FUNCTION_BLOCK IO_RouteDI (* Picks the way an IO block reaches its signal from the Address (a Pi line, a local IO handle, Modbus or simulated) and passes values through that way only. Technical: Backend router for IO_DI; Address: 'gpio[chip:line(:pull_up|:pull_down)(:active_low)]' or 'pwm[chip:channel:period_ns]' a Raspberry Pi's line, set up here; 'modbus[...]' a Modbus CLIENT ID; 'sim' simulated; another name a local IO handle set up elsewhere (IX/QX PARAMS); empty: not connected (QO = FALSE) *)
  (* Standard: 61499-2 *)
  (* Version 0.1, 2026-09-28, Project contributors, AAU Smart Production Lab *)
  PACKAGE modlib;
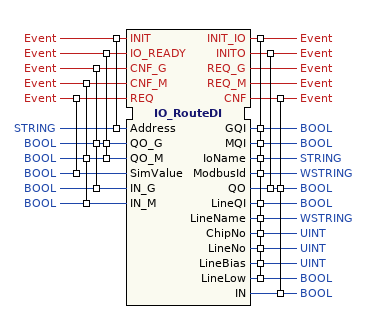
  EVENT_INPUT
    INIT WITH Address; (* Work out from Address how the point is reached *)
    IO_READY WITH QO_G, QO_M; (* The line, the local IO block and the Modbus client are initialised *)
    CNF_G WITH QO_G, IN_G; (* The local IO block answered *)
    CNF_M WITH QO_M, IN_M; (* The Modbus client answered *)
    REQ WITH SimValue; (* Access the point *)
  END_EVENT
  EVENT_OUTPUT
    INIT_IO WITH GQI, MQI, IoName, ModbusId, LineQI, LineName, ChipNo, LineNo, LineBias, LineLow; (* Set up the line, the local IO block and the Modbus client (each only if it is the way) *)
    INITO WITH QO; (* Initialised: QO says whether the point is reachable *)
    REQ_G; (* Access the point through the local IO block (IX/QX/IW/QW) *)
    REQ_M; (* Access the point through the Modbus client *)
    CNF WITH QO, IN; (* Done: QO says whether it worked *)
  END_EVENT
  VAR_INPUT
    Address : STRING; (* Where the point is: 'gpio[chip:line(:pull_up|:pull_down)(:active_low)]', 'pwm[chip:channel:period_ns]', 'modbus[...]', 'sim', or an IO handle's name; empty: not connected *)
    QO_G : BOOL; (* The local IO block works *)
    QO_M : BOOL; (* The Modbus client works *)
    SimValue : BOOL; (* The value read when the address is 'sim' *)
    IN_G : BOOL; (* The raw value read through the local IO block *)
    IN_M : BOOL; (* The raw value read through Modbus *)
  END_VAR
  VAR_OUTPUT
    GQI : BOOL; (* Use the local IO block *)
    MQI : BOOL; (* Use the Modbus client *)
    IoName : STRING; (* The local IO handle's name (PARAMS of IX/QX/IW/QW) *)
    ModbusId : WSTRING; (* The Modbus CLIENT's ID *)
    QO : BOOL; (* The point is reachable, the last access worked *)
    LineQI : BOOL; (* Set up a Raspberry Pi line here (a gpio[...] or pwm[...] address) *)
    LineName : WSTRING; (* The name the line is registered under (the address) *)
    ChipNo : UINT; (* The GPIO or PWM chip's number *)
    LineNo : UINT; (* The GPIO line's or PWM channel's number *)
    LineBias : UINT; (* GPIO bias: 0 none, 2 pull-up, 3 pull-down (FORTE 3.3.0's numbering) *)
    LineLow : BOOL; (* The line is active low *)
    IN : BOOL; (* The value read (an analog one scaled) *)
  END_VAR
  VAR
    Backend : USINT;
  END_VAR
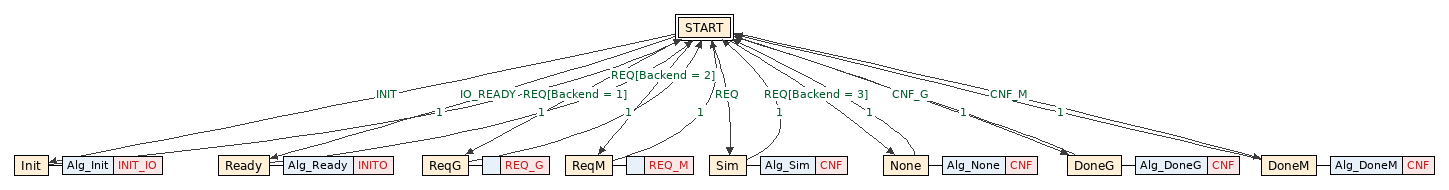
  EC_STATES
    START;
    Init : Alg_Init -> INIT_IO;
    Ready : Alg_Ready -> INITO;
    ReqG : -> REQ_G;
    ReqM : -> REQ_M;
    Sim : Alg_Sim -> CNF;
    None : Alg_None -> CNF;
    DoneG : Alg_DoneG -> CNF;
    DoneM : Alg_DoneM -> CNF;
  END_STATES
  EC_TRANSITIONS
    START TO Init := INIT;
    Init TO START := 1;
    START TO Ready := IO_READY;
    Ready TO START := 1;
    START TO ReqG := REQ[Backend = 1];
    START TO ReqM := REQ[Backend = 2];
    START TO None := REQ[Backend = 3];
    START TO Sim := REQ;
    START TO DoneG := CNF_G;
    START TO DoneM := CNF_M;
    ReqG TO START := 1;
    ReqM TO START := 1;
    Sim TO START := 1;
    None TO START := 1;
    DoneG TO START := 1;
    DoneM TO START := 1;
  END_TRANSITIONS
  ALGORITHM Alg_Init IN ST:
VAR_TEMP
  Field : STRING;
  Length : INT;
  Cut : INT;
  Pos : INT;
  Digit : INT;
  Number : UDINT;
END_VAR
Backend := 3;
LineQI := FALSE;
IF Address = 'sim' THEN
  Backend := 0;
ELSIF LEFT(Address, 7) = 'modbus[' THEN
  Backend := 2;
  ModbusId := STRING_TO_WSTRING(Address);
ELSIF LEFT(Address, 5) = 'gpio[' THEN
  Backend := 1;
  IoName := Address;
  LineQI := TRUE;
  LineName := STRING_TO_WSTRING(Address);
  Length := LEN(Address);
  Field := MID(Address, Length - 5, 6);
  Cut := FIND(Field, ':');
  IF Cut = 0 THEN
    Cut := FIND(Field, ']');
  END_IF;
  Number := 0;
  FOR Digit := 1 TO Cut - 1 DO
    Pos := FIND('0123456789', MID(Field, 1, Digit));
    Number := Number * 10 + INT_TO_UDINT(Pos - 1);
  END_FOR;
  ChipNo := UDINT_TO_UINT(Number);
  Length := LEN(Field);
  Field := MID(Field, Length - Cut, Cut + 1);
  Cut := FIND(Field, ':');
  IF Cut = 0 THEN
    Cut := FIND(Field, ']');
  END_IF;
  Number := 0;
  FOR Digit := 1 TO Cut - 1 DO
    Pos := FIND('0123456789', MID(Field, 1, Digit));
    Number := Number * 10 + INT_TO_UDINT(Pos - 1);
  END_FOR;
  LineNo := UDINT_TO_UINT(Number);
  Length := LEN(Field);
  Field := MID(Field, Length - Cut, Cut + 1);
  IF FIND(Address, ':pull_up') > 0 THEN
    LineBias := 2;
  ELSIF FIND(Address, ':pull_down') > 0 THEN
    LineBias := 3;
  ELSE
    LineBias := 0;
  END_IF;
  LineLow := FIND(Address, ':active_low') > 0;
ELSIF LEN(Address) > 0 THEN
  Backend := 1;
  IoName := Address;
END_IF;
GQI := Backend = 1;
MQI := Backend = 2;
  END_ALGORITHM
  ALGORITHM Alg_Ready IN ST:
QO := (Backend = 0) OR ((Backend = 1) AND QO_G) OR ((Backend = 2) AND QO_M);
  END_ALGORITHM
  ALGORITHM Alg_Sim IN ST:
QO := TRUE;
IN := SimValue;
  END_ALGORITHM
  ALGORITHM Alg_None IN ST:
QO := FALSE;
  END_ALGORITHM
  ALGORITHM Alg_DoneG IN ST:
QO := QO_G;
IN := IN_G;
  END_ALGORITHM
  ALGORITHM Alg_DoneM IN ST:
QO := QO_M;
IN := IN_M;
  END_ALGORITHM
END_FUNCTION_BLOCK
